(* IEC 61131-3 sources: kns-port-domestic/upstream/plc-process-lib/src/Interfaces/I_Alarm, 1 file *)

(* ---- Shelve.method.decl.st ---- *)
// Запрос shelve. TRUE — принято: приоритет <> None, tShelveMax > 0, не OutOfService
METHOD Shelve : BOOL
VAR_INPUT
    tDuration : TIME;   // срок; T#0S — tShelveMax, больше tShelveMax — обрезается
END_VAR
